(*
    Status of FB_FlowMeter.
*)
TYPE ST_FlowStatus EXTENDS ST_StatusBase :
STRUCT
    FrequencyHz : REAL;  // Hz, rising edges of the sensor input during the last second
    FlowRate : REAL;     // Cfg.Factor x FrequencyHz
END_STRUCT
END_TYPE

(* stored: Version 1.1.0.1
   DUT ST_FlowStatus: Id {f90f3807-d193-4984-91f4-1f1741633eec} *)
